(* IEC 61131-3 sources: SortJet_MasterSPS_Aufbau.fbsproj/Device.device.xml.v3^/Plc Logic.plclogic.xml.v3^/Application.application.xml.v3^/10_Schnittstellen, 5 files *)

(* ---- MK_Schnittstelle_Sortjet.gvl ---- *)
(* METADATA
{
	"v3Meta": {
		"objectGuid": "7637b519-9876-476d-bbb2-aba53baea77e"
	}
}
*)
{attribute 'allow_unqualified_access'}
NAMESPACE MK_Schnittstelle_Sortjet
VAR_GLOBAL
//-------------------------------------------------------------------------------------------------
// MASCHINEPARAMETER: SCHNITTSTELLE SORTJET
//-------------------------------------------------------------------------------------------------

  (* Hinweis:
     - Das MMI entscheidet wer Master und wer Slave ist.
       Das MMI, das den Status der Verbundstrecke verwaltet ist der Master!
  *)
  apgMKSchnittstelle_SortJet_Remnant : Schnittstelle_SortJet_ST :=
  (
    bDeaktivieren      := FALSE,                // Station deaktiviert (keine Auftraege, keine Referenzfahrt)
    eSchnittstellenTyp := eSchnittstelle_Master // Rolle der SortJet-SortJet-Schnittstelle (Master/Slave)
  );

END_VAR
END_NAMESPACE

(* ---- MK_Station_401.gvl ---- *)
(* METADATA
{
	"v3Meta": {
		"objectGuid": "b6ce0e10-1e09-4711-a6fa-fa87783967b6"
	}
}
*)
{attribute 'allow_unqualified_access'}
NAMESPACE MK_Station_401
VAR_GLOBAL
//-------------------------------------------------------------------------------------------------
// MASCHINEPARAMETER: SCHNITTSTELLE 401
//-------------------------------------------------------------------------------------------------

  apgMKStation401 : Parameter_Station :=
    (
      stStationsNummern                     := ( NummerIntern    :=   401,                           // Stationsnummer fuer das MMI und die Stationsangabe der Meldungen
                                                 NummerExtern    :=  1401,                           // Stationsnummer fuer Bedienermeldungen
                                                 NummerSPS       :=   401 ),                         // Stationsnummer SPS-intern (Indizes)
      bDeaktivieren                         := TRUE,                                                 // Station deaktiviert (keine Auftraege, keine Referenzfahrt)
      wMeldungsNummer                       := 1300,                                                 // Basis-Meldungsnummer (WatchIO)
      eStationsTyp                          := eFremdanlage,                                         // Typ der Station
      eaAutomatikkreis                      := [eAutomatikkreis_Undefiniert],                        // Automatikkreise, zu denen die Station gehoert
      // stStationsOptionen
      // stStationsAufbau
      // stStationsParameter
      stSchnittstellendaten                 := ( wVorgaengerStation := cSTATION_DEFAULT,             // Station vor dieser Station (cSTATION_DYNAMISCH bei mehreren)
                                                 wNachfolgerStation := cSTATION_DEFAULT,             // Station nach dieser Station (cSTATION_DYNAMISCH bei mehreren)
                                                 bStationIstShuttle := FALSE                         // Station ist ein Shuttle
                                               ),
      stFremdanlage                         := ( bWerteSwappen                          := FALSE,    // Bytes der Auftragsdaten (Lade-ID) und der Empfaenger- Geschwindigkeit swappen
                                                 bCounterSwappen                        := FALSE,    // Nur die bytes von Life Counter swappen
                                                 bSignaleSwappen                        := FALSE,    // Nur die bytes der Signale swappen
                                                 bAnzahlScheibenSwappen                 := FALSE,    // Nur die Bytes der Anzahl Scheiben swappen
                                                 bRemoveETX                             := TRUE,     // ETX aus den Scheiben-IDs des MMI entfernen (Auftragsdaten Fremdanlage)
                                                 tZeitHornAktiv                         := T#5S,     // Signal bei ISO-Line Event
                                                 rAnalogWertVerhaeltniss                := 32.768,   // Umrechnungsfaktor für den Analogwert
                                                 rLaengeStation                         := 0.0,      // Laenge der Fremdanlage (Wegueberwachung der ersten Scheibe in der Nachbarstation), 0 = unbekannt
                                                 wMindestAnalogWert                     := 100,      // Mindestwert, den der Analogwert haben muss um gültig zu sein
                                                 bAnzeigeISOLinieEventAktiv             := FALSE,    // ISO Line Events sollen angezeigt werden
                                                 bAnalogwertAktiv                       := FALSE,    // Geschwindigkeit - Analog | Statische
                                                 rGeschwindigkeit                       := 667,      // Feste Geschwindigkeit der Fremdanlage - (Fester Sollwert)
                                                 rMindestGeschwindigkeitsAenderung      := 5.0,      // Glaettung: Mindestaenderung [mm/s] bevor eine neue Geschwindigkeit uebernommen wird
                                                 tMindestZeitZwischenGeschwAenderung    := T#500MS,  // Glaettung: Mindestzeit zwischen zwei Geschwindigkeitsaenderungen
                                                 rMaxAnalogGeschwindigkeit              := 1000.0,   // Analogwert: Begrenzung der Geschwindigkeit [mm/s]
                                                 eTypSchnittstelle                      := eDefault, // Variante der Schnittstelle
                                                 bStationStatusZuGlasAbruf              := FALSE,    // Stationsstatus beim Glasabruf melden (ISO-Linie)
                                                 bSignaleLoggen                         := TRUE      // Schnittstellensignale loggen
                                               ),
      // stGlasdaten
      eaSicherheitskreis                    := [eSicherheitskreis_Undefiniert],                      // Sicherheitskreise, in die die Station eingebunden ist
      // astSicherheitskreisTeilabschaltung
      eSystemcheckZyklus                    := eSystemcheckZyklus_Undefiniert                        // In welchem Zyklus des Systemchecks die Station geprueft wird
      // astShuttleAnhaltenQuellen
   );

END_VAR
END_NAMESPACE

(* ---- MK_Station_501.gvl ---- *)
(* METADATA
{
	"v3Meta": {
		"objectGuid": "40b5e71b-f854-4565-9b77-acb7772a88ea"
	}
}
*)
{attribute 'allow_unqualified_access'}
NAMESPACE MK_Station_501
VAR_GLOBAL
//-------------------------------------------------------------------------------------------------
// MASCHINEPARAMETER: SCHNITTSTELLE 501
//-------------------------------------------------------------------------------------------------

  apgMKStation501 : Parameter_Station :=
    (
      stStationsNummern                     := ( NummerIntern    :=   501,                           // Stationsnummer fuer das MMI und die Stationsangabe der Meldungen
                                                 NummerExtern    :=  1501,                           // Stationsnummer fuer Bedienermeldungen
                                                 NummerSPS       :=   501 ),                         // Stationsnummer SPS-intern (Indizes)
      bDeaktivieren                         := TRUE,                                                 // Station deaktiviert (keine Auftraege, keine Referenzfahrt)
      wMeldungsNummer                       := 1310,                                                 // Basis-Meldungsnummer (WatchIO)
      eStationsTyp                          := eFremdanlage,                                         // Typ der Station
      eaAutomatikkreis                      := [eAutomatikkreis_Undefiniert],                        // Automatikkreise, zu denen die Station gehoert
      // stStationsOptionen
      // stStationsAufbau
      // stStationsParameter
      stSchnittstellendaten                 := ( wVorgaengerStation := cSTATION_DEFAULT,             // Station vor dieser Station (cSTATION_DYNAMISCH bei mehreren)
                                                 wNachfolgerStation := cSTATION_205,                 // Station nach dieser Station (cSTATION_DYNAMISCH bei mehreren)
                                                 bStationIstShuttle := FALSE                         // Station ist ein Shuttle
                                               ),
      stFremdanlage                         := ( bWerteSwappen                          := FALSE,    // Bytes der Auftragsdaten (Lade-ID) und der Empfaenger- Geschwindigkeit swappen
                                                 bCounterSwappen                        := FALSE,    // Nur die bytes von Life Counter swappen
                                                 bSignaleSwappen                        := FALSE,    // Nur die bytes der Signale swappen
                                                 bAnzahlScheibenSwappen                 := FALSE,    // Nur die Bytes der Anzahl Scheiben swappen
                                                 bRemoveETX                             := TRUE,     // ETX aus den Scheiben-IDs des MMI entfernen (Auftragsdaten Fremdanlage)
                                                 tZeitHornAktiv                         := T#5S,     // Signal bei ISO-Line Event
                                                 rAnalogWertVerhaeltniss                := 32.768,   // Umrechnungsfaktor für den Analogwert
                                                 rLaengeStation                         := 0.0,      // Laenge der Fremdanlage (Wegueberwachung der ersten Scheibe in der Nachbarstation), 0 = unbekannt
                                                 wMindestAnalogWert                     := 100,      // Mindestwert, den der Analogwert haben muss um gültig zu sein
                                                 bAnzeigeISOLinieEventAktiv             := FALSE,    // ISO Line Events sollen angezeigt werden
                                                 bAnalogwertAktiv                       := FALSE,    // Geschwindigkeit - Analog | Statische
                                                 rGeschwindigkeit                       := 350,      // Feste Geschwindigkeit der Fremdanlage - (Fester Sollwert)
                                                 rMindestGeschwindigkeitsAenderung      := 5.0,      // Glaettung: Mindestaenderung [mm/s] bevor eine neue Geschwindigkeit uebernommen wird
                                                 tMindestZeitZwischenGeschwAenderung    := T#500MS,  // Glaettung: Mindestzeit zwischen zwei Geschwindigkeitsaenderungen
                                                 rMaxAnalogGeschwindigkeit              := 1000.0,   // Analogwert: Begrenzung der Geschwindigkeit [mm/s]
                                                 eTypSchnittstelle                      := eDefault, // Variante der Schnittstelle
                                                 bStationStatusZuGlasAbruf              := FALSE,    // Stationsstatus beim Glasabruf melden (ISO-Linie)
                                                 bSignaleLoggen                         := TRUE      // Schnittstellensignale loggen
                                               ),
      // stGlasdaten
      eaSicherheitskreis                    := [eSicherheitskreis_Undefiniert],                      // Sicherheitskreise, in die die Station eingebunden ist
      // astSicherheitskreisTeilabschaltung
      eSystemcheckZyklus                    := eSystemcheckZyklus_Undefiniert                        // In welchem Zyklus des Systemchecks die Station geprueft wird
      // astShuttleAnhaltenQuellen
   );

END_VAR
END_NAMESPACE

(* ---- Konfiguration_Schnittstelle_401.gvl ---- *)
(* METADATA
{
	"v3Meta": {
		"objectGuid": "8cc29e57-f99b-4de6-9b97-bbeab92ab639"
	}
}
*)
{attribute 'allow_unqualified_access'}
NAMESPACE Konfiguration_Schnittstelle_401
VAR_CONFIG

//-------------------------------------------------------------------------------------------------
// KONFIGURATION: SCHNITTSTELLE 401 Auslauf Glaston mit Koppler
//-------------------------------------------------------------------------------------------------
  // ------------------------------------ HARDWARE EINGAENGE ---------------------------------------
  // Standard Eingaenge
  Globale_Bausteine.aSchnittstelleAuslauf[401].in_bTasterGlasbruch                          AT %MX1.0    : BOOL; // OPTION
  Globale_Bausteine.aSchnittstelleAuslauf[401].in_bTasterSpezial                            AT %MX1.0    : BOOL; // OPTION
  // Koppler Eingaenge (Empfaenger -> Sender)
  Globale_Bausteine.aSchnittstelleAuslauf[401].in_wEmpfaengerLiveCounter                    AT %MW100    : WORD; // OPTION - Wort 0 LiveCounter gespiegelt
  Globale_Bausteine.aSchnittstelleAuslauf[401].in_awEmpfaengerLadeIDGespiegelt              AT %MW100    : ARRAY [1..8] OF WORD; // OPTION - Wort 1..8 Lade-ID gespiegelt
  Globale_Bausteine.aSchnittstelleAuslauf[401].in_wEmpfaengerSignale                        AT %MW100    : WORD; // OPTION - Wort 49 Signale
  Globale_Bausteine.aSchnittstelleAuslauf[401].in_dwEmpfaengerGeschwindigkeit               AT %MD50     : DWORD; // OPTION - Wort 50 Geschwindigkeit [mm/s]
  Globale_Bausteine.aSchnittstelleAuslauf[401].in_wEmpfaengerRampe                          AT %MW100    : WORD; // OPTION - Wort 52 Rampe [mm/s2]

  // ------------------------------------ HARDWARE AUSGAENGE ---------------------------------------
  // Standard Ausgaenge
  Globale_Bausteine.aSchnittstelleAuslauf[401].out_bSenderBereit                            AT %MX4010.0 : BOOL; // OPTION
  Globale_Bausteine.aSchnittstelleAuslauf[401].out_bSenderGlasBereit                        AT %MX4010.1 : BOOL; // OPTION
  Globale_Bausteine.aSchnittstelleAuslauf[401].out_bLeuchteGlasbruch                        AT %MX4010.2 : BOOL; // OPTION
  Globale_Bausteine.aSchnittstelleAuslauf[401].out_bLeuchteSpezial                          AT %MX4010.3 : BOOL; // OPTION
  Globale_Bausteine.aSchnittstelleAuslauf[401].out_bAmpelEventAktiv                         AT %MX4010.4 : BOOL; // OPTION
  Globale_Bausteine.aSchnittstelleAuslauf[401].Horn.out_bHorn                               AT %MX4010.5 : BOOL; // OPTION
  // Koppler Ausgaenge (Sender -> Empfaenger)
  Globale_Bausteine.aSchnittstelleAuslauf[401].out_wSenderLiveCounter                       AT %MW4010   : WORD; // OPTION - Wort 0 LiveCounter
  Globale_Bausteine.aSchnittstelleAuslauf[401].out_wSenderSignale                           AT %MW4011   : WORD; // OPTION - Wort 50 Signale
  Globale_Bausteine.aSchnittstelleAuslauf[401].out_awSenderLadeID                           AT %MW4012   : ARRAY [1..8] OF WORD; // OPTION - Wort 1..8 Lade-ID (%MW4012..%MW4019)

END_VAR

END_NAMESPACE

(* ---- Konfiguration_Schnittstelle_501.gvl ---- *)
(* METADATA
{
	"v3Meta": {
		"objectGuid": "64e1a0cc-c108-4526-a679-59adff7e9323"
	}
}
*)
{attribute 'allow_unqualified_access'}
NAMESPACE Konfiguration_Schnittstelle_501
VAR_CONFIG

//-------------------------------------------------------------------------------------------------
// KONFIGURATION: SCHNITTSTELLE 501 Einlauf VSG (Station 205)
//-------------------------------------------------------------------------------------------------
  // ------------------------------------ HARDWARE EINGAENGE ---------------------------------------
  // Standard Eingaenge
  Globale_Bausteine.aSchnittstelleEinlauf[501].in_bTasterGlasbruch                          AT %IX9.5    : BOOL; // IO-L - Signal 1 von VSG
  Globale_Bausteine.aSchnittstelleEinlauf[501].in_bTasterSpezial                            AT %IX9.6    : BOOL; // IO-L - Signal 2 von VSG
  // VSG Eingaenge
  Globale_Bausteine.aSchnittstelleEinlauf[501].in_bAutomatikBetrieb                         AT %IX9.7    : BOOL; // IO-L - Signal 3 von VSG (VSG im Automatikbetrieb)
  Globale_Bausteine.aSchnittstelleEinlauf[501].in_bGlasBereit                               AT %IX10.0   : BOOL; // IO-L - Signal 4 von VSG (VSG Glas bereit)

  // ------------------------------------ HARDWARE AUSGAENGE ---------------------------------------
  // Standard Ausgaenge
  Globale_Bausteine.aSchnittstelleEinlauf[501].out_bSenderBereit                            AT %QX7.3    : BOOL; // IO-L - Signal 5 an VSG
  Globale_Bausteine.aSchnittstelleEinlauf[501].out_bSenderGlasBereit                        AT %QX7.4    : BOOL; // IO-L - Signal 6 an VSG
  Globale_Bausteine.aSchnittstelleEinlauf[501].out_bLeuchteGlasbruch                        AT %QX7.5    : BOOL; // IO-L - Signal 7 an VSG
  Globale_Bausteine.aSchnittstelleEinlauf[501].out_bLeuchteSpezial                          AT %QX7.6    : BOOL; // IO-L - Signal 8 an VSG
  Globale_Bausteine.aSchnittstelleEinlauf[501].out_bAmpelEventAktiv                         AT %MX5010.4 : BOOL; // OPTION
  Globale_Bausteine.aSchnittstelleEinlauf[501].Horn.out_bHorn                               AT %MX5010.5 : BOOL; // OPTION
  // VSG Ausgaenge
  Globale_Bausteine.aSchnittstelleEinlauf[501].out_bEinlaufsensor                           AT %MX5010.6 : BOOL; // OPTION - Einlaufsensor an VSG
  Globale_Bausteine.aSchnittstelleEinlauf[501].out_bBereitZumEintrasport                    AT %MX5010.7 : BOOL; // OPTION - bereit zum Eintransport

END_VAR

END_NAMESPACE
